// TIA Portal V19 export
// export: Created 2026-10-15T10:10:35.541158Z, ExportSetting WithDefaults, DisplayName Totally Integrated Automation Portal, DisplayVersion V19, DisplayName TIA Portal Openness, DisplayVersion V19, DisplayName TIA Portal Version Control Interface, DisplayVersion V19, DisplayName STEP 7 Professional, DisplayVersion V19, DisplayName STEP 7 Safety, DisplayVersion V19, DisplayName WinCC Basic/Comfort/Advanced, DisplayVersion V19, DisplayName WinCC Unified, DisplayVersion V19
FUNCTION "ROLL_PB8" : Void   // FC18, SCL
{ S7_Optimized_Access := 'TRUE' }
VERSION : 0.1
// stored: AutoNumber true, IsIECCheckEnabled false, SetENOAutomatically false, UDAEnableTagReadback false
   VAR_TEMP
      r : Bool;
      a1 : Word;
      a2 : Word;
      activeDataBlock : Int;
      comparisonResults : Array[0..0] of Bool;
   END_VAR
BEGIN

   #r := FALSE;
   #a1 := W#16#0000;
   #a2 := W#16#0000;
   #activeDataBlock := 0;
   // PB8, STEP 5 network 1
   #r := ("ROLL_State".M[37, 7] OR "ROLL_State".M[38, 0] OR "ROLL_State".M[39, 7] OR "ROLL_State".M[40, 0] OR "ROLL_State".M[40, 1] OR "ROLL_State".M[40, 4] OR "ROLL_State".M[41, 0] OR "ROLL_State".M[41, 6] OR "ROLL_State".M[41, 7] OR "ROLL_State".M[42, 2] OR "ROLL_State".M[42, 3]);
   "ROLL_State".M[33, 0] := #r;
   // PB8, STEP 5 network 2
   #r := (((NOT "ROLL_State".M[16, 0]) AND (NOT "ROLL_State".M[16, 1]) AND (NOT "ROLL_State".M[16, 4]) AND "ROLL_State".M[37, 2]) OR "ROLL_State".M[37, 3] OR "ROLL_State".M[37, 5] OR "ROLL_State".M[37, 6] OR "ROLL_State".M[39, 4] OR "ROLL_State".M[39, 5] OR "ROLL_State".M[40, 2] OR "ROLL_State".M[40, 3] OR "ROLL_State".M[40, 6] OR "ROLL_State".M[40, 7] OR "ROLL_State".M[41, 2] OR "ROLL_State".M[42, 0] OR "ROLL_State".M[42, 4]);
   "ROLL_State".M[33, 1] := #r;
   // PB8, STEP 5 network 3
   #a2 := #a1;
   #a1 := W#16#2030;
   #r := ((NOT "ROLL_State".M[3, 1]) AND ("ROLL_State".M[33, 0] OR "ROLL_State".M[42, 6] OR "ROLL_State".M[43, 4] OR "ROLL_State".M[43, 6] OR "ROLL_State".M[43, 7] OR "ROLL_State".M[44, 2] OR "ROLL_State".M[45, 0] OR "ROLL_State".M[45, 1] OR "ROLL_State".M[45, 5] OR "ROLL_State".M[45, 7] OR "ROLL_State".M[46, 1] OR "ROLL_State".M[46, 4] OR "ROLL_State".M[46, 6] OR "ROLL_State".M[52, 1] OR "ROLL_State".M[52, 2] OR "ROLL_State".M[53, 3]) AND "ROLL_IO".Input[0, 2] AND "ROLL_State".M[29, 0]);
   "ROLL_TimerOp"(Number := 40,
                  Operation := 0,
                  Signal := #r,
                  Preset := #a1);
   // PB8, STEP 5 network 4
   #a2 := #a1;
   #a1 := W#16#2030;
   #r := ((NOT "ROLL_State".M[3, 1]) AND (((NOT "ROLL_IO".Input[11, 2]) AND "ROLL_State".M[52, 0]) OR ((NOT "ROLL_State".M[15, 1]) AND "ROLL_State".M[53, 1]) OR "ROLL_State".M[33, 1] OR "ROLL_State".M[43, 0] OR "ROLL_State".M[43, 2] OR "ROLL_State".M[43, 3] OR "ROLL_State".M[44, 0] OR "ROLL_State".M[44, 7] OR "ROLL_State".M[45, 3] OR "ROLL_State".M[45, 4] OR "ROLL_State".M[46, 2] OR "ROLL_State".M[46, 3] OR "ROLL_State".M[46, 7] OR "ROLL_State".M[47, 3] OR "ROLL_State".M[52, 3] OR "ROLL_State".M[53, 2] OR "ROLL_State".M[53, 5] OR "ROLL_State".M[53, 6]) AND "ROLL_IO".Input[0, 2] AND "ROLL_State".M[29, 0]);
   "ROLL_TimerOp"(Number := 41,
                  Operation := 0,
                  Signal := #r,
                  Preset := #a1);
   // PB8, STEP 5 network 5
   #r := ("ROLL_State".S5Timers[40].Q OR "ROLL_State".S5Timers[41].Q);
   IF #r THEN
       "ROLL_State".M[34, 1] := TRUE;
   END_IF;
   #r := ((NOT "ROLL_IO".Input[0, 2]) OR "ROLL_State".M[3, 1]);
   IF #r THEN
       "ROLL_State".M[34, 1] := FALSE;
   END_IF;
   // PB8, STEP 5 network 6
   RETURN;
END_FUNCTION
